(* IEC 61131-3 sources: SemantiST/compiler/intake/normalize/probes/scl-quoted-identifier, 2 files *)

(* ---- original.st ---- *)
FUNCTION "Scale Value" : INT
VAR_INPUT
    X : INT;
END_VAR
"Scale Value" := X * 5;
END_FUNCTION

FUNCTION main : DINT
printf('%d$N', "Scale Value"(3));
main := 0;
END_FUNCTION

(* ---- rewritten.st ---- *)
FUNCTION Scale_Value__Q : INT
VAR_INPUT
    X : INT;
END_VAR
Scale_Value__Q := X * 5;
END_FUNCTION

FUNCTION main : DINT
printf('%d$N', Scale_Value__Q(3));
main := 0;
END_FUNCTION
